// LS Electric XG5000 project: first-out
// PLC LSPLC

PROGRAM first-out (task: 스캔 프로그램)

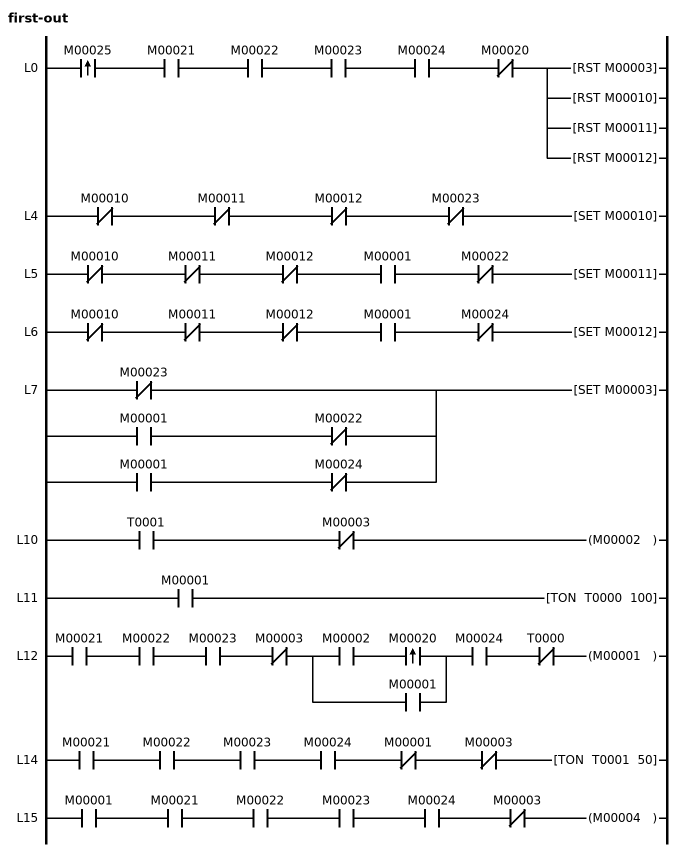
; L0
LOADP     M00025
AND       M00021
AND       M00022
AND       M00023
AND       M00024
AND NOT   M00020
RST       M00003
RST       M00010
RST       M00011
RST       M00012
; L4
LOAD NOT  M00010
AND NOT   M00011
AND NOT   M00012
AND NOT   M00023
SET       M00010
; L5
LOAD NOT  M00010
AND NOT   M00011
AND NOT   M00012
AND       M00001
AND NOT   M00022
SET       M00011
; L6
LOAD NOT  M00010
AND NOT   M00011
AND NOT   M00012
AND       M00001
AND NOT   M00024
SET       M00012
; L7
LOAD NOT  M00023
LOAD      M00001
AND NOT   M00022
OR LOAD
LOAD      M00001
AND NOT   M00024
OR LOAD
SET       M00003
; L10
LOAD      T0001
AND NOT   M00003
OUT       M00002
; L11
LOAD      M00001
TON       T0000 100
; L12
LOAD      M00021
AND       M00022
AND       M00023
AND NOT   M00003
LOAD      M00002
ANDP      M00020
OR        M00001
AND LOAD
AND       M00024
AND NOT   T0000
OUT       M00001
; L14
LOAD      M00021
AND       M00022
AND       M00023
AND       M00024
AND NOT   M00001
AND NOT   M00003
TON       T0001 50
; L15
LOAD      M00001
AND       M00021
AND       M00022
AND       M00023
AND       M00024
AND NOT   M00003
OUT       M00004